FUNCTION_BLOCK EquipmentGroup IMPLEMENTS I_Diagnosable, I_Resettable
VAR CONSTANT
    MaxChildren : DINT := 16;
END_VAR
VAR
    _Name        : STRING(32);
    _Children    : ARRAY[0..MaxChildren - 1] OF I_Diagnosable;
    _Resettables : ARRAY[0..MaxChildren - 1] OF I_Resettable;
    _Count       : DINT;
END_VAR
(*
    EquipmentGroup

    A named group of devices or other groups, behind the same interfaces
    as one device. It has a fault while any child has one, and reports
    the first faulted child's text, prefixed with that child's name.
    Reset() resets every child that implements I_Resettable.
    AddChild() is called while wiring, before the group is first asked.
*)

METHOD FB_init : BOOL
VAR_INPUT
    bInitRetains : BOOL;
    bInCopyCode  : BOOL;
    Name         : STRING(32);
END_VAR
_Name := Name;
END_METHOD

METHOD PUBLIC AddChild : BOOL
VAR_INPUT
    Child : I_Diagnosable;
END_VAR
VAR
    Me         : I_Diagnosable;
    Resettable : I_Resettable;
    i          : DINT;
END_VAR
Me := THIS^;
IF Child = 0 OR Child = Me OR _Count >= MaxChildren THEN
    AddChild := FALSE;
    RETURN;
END_IF
FOR i := 0 TO _Count - 1 DO           // the same child only once
    IF _Children[i] = Child THEN
        AddChild := FALSE;
        RETURN;
    END_IF
END_FOR
_Children[_Count] := Child;
IF __QUERYINTERFACE(Child, Resettable) THEN
    _Resettables[_Count] := Resettable;
END_IF
_Count := _Count + 1;
AddChild := TRUE;
END_METHOD

METHOD PUBLIC Reset
VAR
    i : DINT;
END_VAR
FOR i := 0 TO _Count - 1 DO
    IF _Resettables[i] <> 0 THEN
        _Resettables[i].Reset();
    END_IF
END_FOR
END_METHOD

METHOD PRIVATE FirstFaultIndex : DINT
VAR
    i : DINT;
END_VAR
FOR i := 0 TO _Count - 1 DO
    IF _Children[i].HasFault THEN
        FirstFaultIndex := i;
        RETURN;
    END_IF
END_FOR
FirstFaultIndex := _Count;            // no child has a fault
END_METHOD

METHOD PRIVATE DescribeFault : STRING
VAR_INPUT
    Index : DINT;
END_VAR
IF Index < _Count THEN
    DescribeFault := CONCAT(CONCAT(_Children[Index].Name, ': '), _Children[Index].FaultText);
END_IF
END_METHOD

PROPERTY PUBLIC Name : STRING
GET
Name := _Name;
END_GET
END_PROPERTY

PROPERTY PUBLIC HasFault : BOOL
GET
HasFault := FirstFaultIndex() < _Count;
END_GET
END_PROPERTY

PROPERTY PUBLIC FaultText : STRING
GET
FaultText := DescribeFault(Index := FirstFaultIndex());
END_GET
END_PROPERTY

PROPERTY PUBLIC ChildCount : DINT
GET
ChildCount := _Count;
END_GET
END_PROPERTY

END_FUNCTION_BLOCK

(* stored: Version 1.1.0.1, ProductVersion 3.1.4026.0
   POU EquipmentGroup: Id {df4d33af-2551-433b-8607-e9e14ad03a2e}, SpecialFunc None
   Folder I_Diagnosable: Id {dbc7c784-3082-4e7a-a527-52be38b83f31}
   Folder I_Resettable: Id {5b93e3e1-9ead-48ca-b8de-caa4b189f039}
   Method FB_init: Id {37459d52-9f7c-4e5c-80cd-c895d42c7ab4}
   Method AddChild: Id {2abd6778-5a9d-480f-a4d1-978c85c747ec}
   Method Reset: Id {d83eb1a0-a4bb-4045-a892-564ca39b5da8}
   Method FirstFaultIndex: Id {f829a151-4e73-404f-9013-ffc49c6a383e}
   Method DescribeFault: Id {e73c7bb2-f2f3-431d-85ed-7dea1d468da0}
   Property Name: Id {7aa0ad69-5184-4be1-bb25-58f4f5070a4f}
   Get Get: Id {bbf64da4-f5f9-4a9c-b080-4edd5a761c2b}
   Property HasFault: Id {191cd794-1cc7-4833-bb2d-a4c912d04755}
   Get Get: Id {2c5f48dd-947e-4748-b9ee-6a95ad8d84df}
   Property FaultText: Id {81bdde44-aee3-46a5-bfae-3cca9fe62f90}
   Get Get: Id {5c8f35b8-cc50-4198-b37e-64ded9a506b5}
   Property ChildCount: Id {22bb6ff0-1add-4a6f-bcf2-87e79716d8fa}
   Get Get: Id {dea68905-fd9c-479d-88e3-0a4d2d5137b5} *)
